// TIA Portal V21 export
// export: Created 2026-08-21T20:18:56.8121563Z, ExportSetting None, DisplayName Totally Integrated Automation Portal, DisplayVersion V21, DisplayName STEP 7 Professional, DisplayVersion V21, DisplayName STEP 7 Safety, DisplayVersion V21, DisplayName Tech WebApplication, DisplayVersion V21, DisplayName WinCC Basic/Comfort/Advanced, DisplayVersion V21, DisplayName WinCC Professional, DisplayVersion V21, DisplayName WinCC Unified, DisplayVersion V21
TYPE "UDT_Service_StepRawDataMedium"
   STRUCT
      "step" : Array[0..99] of "UDT_Service_StepMedium";
      parameterDefinition : Array[0..31] of "UDT_Service_ParameterDefinition";
   END_STRUCT;
END_TYPE
